Fanuc KAREL source: kb00024.KL

-- PROVISIONAL review KL for V1013-1; original PC SHA256 de674383d34266390a8aa9e5e7be8dd5abc7eb85d058e7025d586c5407dc1950
-- Incomplete behavior may be omitted. Consult companion uncertainty JSON. Do not deploy.
PROGRAM KB00024
%NOLOCKGROUP
BEGIN
  -- UNRESOLVED_PC offsets 5-15; opcodes 27,22,31
  -- UNRESOLVED_PC offsets 20-24; opcodes 7F
END KB00024
